PROGRAM MAIN
VAR
    bReady : BOOL := TRUE;
END_VAR

END_PROGRAM

(* stored: Version 1.1.0.1
   POU MAIN: Id {26bcb203-7e0c-455c-9b18-2b2b483f83c4}, SpecialFunc None *)
